// TIA Portal V20 export
Screen "Andon"  1276x673
  ScreenItem "Title_ScreenOverview_X390_Y2" at 9,7 size 1265x44  Type=HmiTextBox
  ScreenItem "permanentareaborderrectangle" at 0,0 size 0x0  Type=HmiRectangle
  ScreenItem "Text box_3" at 346,188 size 590x89  Type=HmiTextBox
  ScreenItem "Title_ScreenOverview_X390_Y2_1" at 9,97 size 84x44  Type=HmiTextBox
  ScreenItem "IO 域_19" at 9,142 size 84x44  Type=HmiIOField
  ScreenItem "Title_ScreenOverview_X390_Y2_5" at 261,97 size 84x44  Type=HmiTextBox
  ScreenItem "IO 域_21" at 261,142 size 84x44  Type=HmiIOField
  ScreenItem "Title_ScreenOverview_X390_Y2_3" at 93,97 size 84x44  Type=HmiTextBox
  ScreenItem "IO 域_5" at 93,142 size 84x44  Type=HmiIOField
  ScreenItem "Title_ScreenOverview_X390_Y2_4" at 177,97 size 84x44  Type=HmiTextBox
  ScreenItem "IO 域_20" at 177,142 size 84x44  Type=HmiIOField
  ScreenItem "Title_ScreenOverview_X390_Y2_6" at 345,97 size 84x44  Type=HmiTextBox
  ScreenItem "IO 域_22" at 345,142 size 84x44  Type=HmiIOField
  ScreenItem "Title_ScreenOverview_X390_Y2_11" at 9,52 size 252x44  Type=HmiTextBox
  ScreenItem "Title_ScreenOverview_X390_Y2_18" at 431,97 size 84x44  Type=HmiTextBox
  ScreenItem "IO 域_42" at 431,142 size 84x44  Type=HmiIOField
  ScreenItem "Title_ScreenOverview_X390_Y2_19" at 683,97 size 84x44  Type=HmiTextBox
  ScreenItem "IO 域_43" at 683,142 size 84x44  Type=HmiIOField
  ScreenItem "Title_ScreenOverview_X390_Y2_20" at 515,97 size 84x44  Type=HmiTextBox
  ScreenItem "IO 域_44" at 515,142 size 84x44  Type=HmiIOField
  ScreenItem "Title_ScreenOverview_X390_Y2_21" at 599,97 size 84x44  Type=HmiTextBox
  ScreenItem "IO 域_45" at 599,142 size 84x44  Type=HmiIOField
  ScreenItem "Title_ScreenOverview_X390_Y2_22" at 767,97 size 84x44  Type=HmiTextBox
  ScreenItem "IO 域_46" at 767,142 size 84x44  Type=HmiIOField
  ScreenItem "Title_ScreenOverview_X390_Y2_23" at 431,52 size 252x44  Type=HmiTextBox
  ScreenItem "Title_ScreenOverview_X390_Y2_25" at 1105,97 size 84x44  Type=HmiTextBox
  ScreenItem "IO 域_48" at 1105,142 size 84x44  Type=HmiIOField
  ScreenItem "Title_ScreenOverview_X390_Y2_28" at 1189,97 size 84x44  Type=HmiTextBox
  ScreenItem "IO 域_51" at 1189,142 size 84x44  Type=HmiIOField
  ScreenItem "Title_ScreenOverview_X390_Y2_29" at 853,52 size 252x44  Type=HmiTextBox
  ScreenItem "Title_ScreenOverview_X390_Y2_7" at 9,188 size 84x44  Type=HmiTextBox
  ScreenItem "IO 域_23" at 9,233 size 84x44  Type=HmiIOField
  ScreenItem "Title_ScreenOverview_X390_Y2_8" at 177,188 size 84x44  Type=HmiTextBox
  ScreenItem "IO 域_24" at 177,233 size 84x44  Type=HmiIOField
  ScreenItem "Text box_32" at 262,278 size 255x96  Type=HmiTextBox
  ScreenItem "Text box_33" at 514,278 size 255x96  Type=HmiTextBox
  ScreenItem "Text box_34" at 764,278 size 255x96  Type=HmiTextBox
  ScreenItem "Text box_35" at 1017,278 size 255x96  Type=HmiTextBox
  ScreenItem "Text box_36" at 10,373 size 255x96  Type=HmiTextBox
  ScreenItem "Text box_37" at 262,373 size 255x96  Type=HmiTextBox
  ScreenItem "Title_ScreenOverview_X390_Y2_38" at 93,188 size 84x44  Type=HmiTextBox
  ScreenItem "IO 域_6" at 93,233 size 84x44  Type=HmiIOField
  ScreenItem "Title_ScreenOverview_X390_Y2_39" at 261,188 size 84x44  Type=HmiTextBox
  ScreenItem "IO 域_7" at 261,233 size 84x44  Type=HmiIOField
  ScreenItem "Title_ScreenOverview_X390_Y2_24" at 853,97 size 84x44  Type=HmiTextBox
  ScreenItem "IO 域_47" at 853,142 size 84x44  Type=HmiIOField
  ScreenItem "Title_ScreenOverview_X390_Y2_26" at 937,97 size 84x44  Type=HmiTextBox
  ScreenItem "IO 域_49" at 937,142 size 84x44  Type=HmiIOField
  ScreenItem "Title_ScreenOverview_X390_Y2_27" at 1021,97 size 84x44  Type=HmiTextBox
  ScreenItem "IO 域_50" at 1021,142 size 84x44  Type=HmiIOField
  ScreenItem "Title_ScreenOverview_X390_Y2_9" at 937,188 size 84x44  Type=HmiTextBox
  ScreenItem "IO 域_8" at 937,233 size 84x44  Type=HmiIOField
  ScreenItem "Title_ScreenOverview_X390_Y2_10" at 1021,188 size 84x44  Type=HmiTextBox
  ScreenItem "IO 域_9" at 1021,233 size 84x44  Type=HmiIOField
  ScreenItem "Title_ScreenOverview_X390_Y2_14" at 1105,188 size 84x44  Type=HmiTextBox
  ScreenItem "IO 域_10" at 1105,233 size 84x44  Type=HmiIOField
  ScreenItem "Move_Legend" at 1182,7 size 90x44  Type=HmiButton
  ScreenItem "Title_ScreenOverview_X390_Y2_17" at 1189,188 size 84x44  Type=HmiTextBox
  ScreenItem "IO 域_11" at 1189,233 size 84x44  Type=HmiIOField
  ScreenItem "IO field_1" at 9,7 size 168x44  Type=HmiIOField
  ScreenItem "Title_ScreenOverview_X390_Y2_13" at 262,52 size 84x44  Type=HmiTextBox
  ScreenItem "IO 域_12" at 346,52 size 84x44  Type=HmiIOField
  ScreenItem "IO 域_13" at 767,52 size 84x44  Type=HmiIOField
  ScreenItem "Title_ScreenOverview_X390_Y2_15" at 683,52 size 84x44  Type=HmiTextBox
  ScreenItem "IO 域_14" at 1188,53 size 84x44  Type=HmiIOField
  ScreenItem "Title_ScreenOverview_X390_Y2_16" at 1104,53 size 84x44  Type=HmiTextBox
  ScreenItem "IO 域_2" at 504,31 size 126x32  Type=HmiIOField
  ScreenItem "Title_ScreenOverview_X390_Y2_31" at 0,31 size 184x32  Type=HmiTextBox
  ScreenItem "IO 域_4" at 185,31 size 126x32  Type=HmiIOField
  ScreenItem "Title_ScreenOverview_X390_Y2_2" at 0,0 size 630x30  Type=HmiTextBox
  ScreenItem "Title_ScreenOverview_X390_Y2_12" at 313,31 size 189x32  Type=HmiTextBox
  ScreenItem "Title_ScreenOverview_X390_Y2_32" at 0,64 size 184x32  Type=HmiTextBox
  ScreenItem "IO 域_3" at 185,64 size 126x32  Type=HmiIOField
  ScreenItem "Title_ScreenOverview_X390_Y2_30" at 313,64 size 189x32  Type=HmiTextBox
  ScreenItem "IO 域_1" at 504,64 size 126x32  Type=HmiIOField
  ScreenItem "IO 域_57" at 1136,31 size 126x32  Type=HmiIOField
  ScreenItem "Title_ScreenOverview_X390_Y2_33" at 632,31 size 184x32  Type=HmiTextBox
  ScreenItem "IO 域_56" at 817,31 size 126x32  Type=HmiIOField
  ScreenItem "Title_ScreenOverview_X390_Y2_34" at 632,0 size 630x30  Type=HmiTextBox
  ScreenItem "Title_ScreenOverview_X390_Y2_35" at 945,31 size 189x32  Type=HmiTextBox
  ScreenItem "Title_ScreenOverview_X390_Y2_36" at 632,64 size 184x32  Type=HmiTextBox
  ScreenItem "IO 域_58" at 817,64 size 126x32  Type=HmiIOField
  ScreenItem "Title_ScreenOverview_X390_Y2_37" at 945,64 size 189x32  Type=HmiTextBox
  ScreenItem "IO 域_59" at 1136,64 size 126x32  Type=HmiIOField
  ScreenItem "IO 域_37" at 504,31 size 126x32  Type=HmiIOField
  ScreenItem "Title_ScreenOverview_X390_Y2_68" at 0,31 size 184x32  Type=HmiTextBox
  ScreenItem "IO 域_53" at 185,31 size 126x32  Type=HmiIOField
  ScreenItem "Title_ScreenOverview_X390_Y2_67" at 0,0 size 630x30  Type=HmiTextBox
  ScreenItem "Title_ScreenOverview_X390_Y2_66" at 313,31 size 189x32  Type=HmiTextBox
  ScreenItem "Title_ScreenOverview_X390_Y2_65" at 0,64 size 184x32  Type=HmiTextBox
  ScreenItem "IO 域_52" at 185,64 size 126x32  Type=HmiIOField
  ScreenItem "Title_ScreenOverview_X390_Y2_64" at 313,64 size 189x32  Type=HmiTextBox
  ScreenItem "IO 域_41" at 504,64 size 126x32  Type=HmiIOField
  ScreenItem "IO 域_40" at 1136,31 size 126x32  Type=HmiIOField
  ScreenItem "Title_ScreenOverview_X390_Y2_63" at 632,31 size 184x32  Type=HmiTextBox
  ScreenItem "IO 域_39" at 817,31 size 126x32  Type=HmiIOField
  ScreenItem "Title_ScreenOverview_X390_Y2_62" at 632,0 size 630x30  Type=HmiTextBox
  ScreenItem "Title_ScreenOverview_X390_Y2_61" at 945,31 size 189x32  Type=HmiTextBox
  ScreenItem "Title_ScreenOverview_X390_Y2_60" at 632,64 size 184x32  Type=HmiTextBox
  ScreenItem "IO 域_38" at 817,64 size 126x32  Type=HmiIOField
  ScreenItem "Title_ScreenOverview_X390_Y2_69" at 945,64 size 189x32  Type=HmiTextBox
  ScreenItem "IO 域_54" at 1136,64 size 126x32  Type=HmiIOField
  ScreenItem "IO 域_15" at 504,31 size 126x32  Type=HmiIOField
  ScreenItem "Title_ScreenOverview_X390_Y2_48" at 0,31 size 184x32  Type=HmiTextBox
  ScreenItem "IO 域_27" at 185,31 size 126x32  Type=HmiIOField
  ScreenItem "Title_ScreenOverview_X390_Y2_47" at 0,0 size 630x30  Type=HmiTextBox
  ScreenItem "Title_ScreenOverview_X390_Y2_46" at 313,31 size 189x32  Type=HmiTextBox
  ScreenItem "Title_ScreenOverview_X390_Y2_45" at 0,64 size 184x32  Type=HmiTextBox
  ScreenItem "IO 域_26" at 185,64 size 126x32  Type=HmiIOField
  ScreenItem "Title_ScreenOverview_X390_Y2_44" at 313,64 size 189x32  Type=HmiTextBox
  ScreenItem "IO 域_25" at 504,64 size 126x32  Type=HmiIOField
  ScreenItem "IO 域_18" at 1136,31 size 126x32  Type=HmiIOField
  ScreenItem "Title_ScreenOverview_X390_Y2_43" at 632,31 size 184x32  Type=HmiTextBox
  ScreenItem "IO 域_17" at 817,31 size 126x32  Type=HmiIOField
  ScreenItem "Title_ScreenOverview_X390_Y2_42" at 632,0 size 630x30  Type=HmiTextBox
  ScreenItem "Title_ScreenOverview_X390_Y2_41" at 945,31 size 189x32  Type=HmiTextBox
  ScreenItem "Title_ScreenOverview_X390_Y2_40" at 632,64 size 184x32  Type=HmiTextBox
  ScreenItem "IO 域_16" at 817,64 size 126x32  Type=HmiIOField
  ScreenItem "Title_ScreenOverview_X390_Y2_49" at 945,64 size 189x32  Type=HmiTextBox
  ScreenItem "IO 域_28" at 1136,64 size 126x32  Type=HmiIOField
  ScreenItem "IO 域_29" at 504,31 size 126x32  Type=HmiIOField
  ScreenItem "Title_ScreenOverview_X390_Y2_58" at 0,31 size 184x32  Type=HmiTextBox
  ScreenItem "IO 域_35" at 185,31 size 126x32  Type=HmiIOField
  ScreenItem "Title_ScreenOverview_X390_Y2_57" at 0,0 size 630x30  Type=HmiTextBox
  ScreenItem "Title_ScreenOverview_X390_Y2_56" at 313,31 size 189x32  Type=HmiTextBox
  ScreenItem "Title_ScreenOverview_X390_Y2_55" at 0,64 size 184x32  Type=HmiTextBox
  ScreenItem "IO 域_34" at 185,64 size 126x32  Type=HmiIOField
  ScreenItem "Title_ScreenOverview_X390_Y2_54" at 313,64 size 189x32  Type=HmiTextBox
  ScreenItem "IO 域_33" at 504,64 size 126x32  Type=HmiIOField
  ScreenItem "IO 域_32" at 1136,31 size 126x32  Type=HmiIOField
  ScreenItem "Title_ScreenOverview_X390_Y2_53" at 632,31 size 184x32  Type=HmiTextBox
  ScreenItem "IO 域_31" at 817,31 size 126x32  Type=HmiIOField
  ScreenItem "Title_ScreenOverview_X390_Y2_52" at 632,0 size 630x30  Type=HmiTextBox
  ScreenItem "Title_ScreenOverview_X390_Y2_51" at 945,31 size 189x32  Type=HmiTextBox
  ScreenItem "Title_ScreenOverview_X390_Y2_50" at 632,64 size 184x32  Type=HmiTextBox
  ScreenItem "IO 域_30" at 817,64 size 126x32  Type=HmiIOField
  ScreenItem "Title_ScreenOverview_X390_Y2_59" at 945,64 size 189x32  Type=HmiTextBox
  ScreenItem "IO 域_36" at 1136,64 size 126x32  Type=HmiIOField
  ScreenItem "Text box_1" at 514,373 size 255x96  Type=HmiTextBox
  ScreenItem "Text box_2" at 10,278 size 255x96  Type=HmiTextBox
  ScreenItem "Text box_4" at 764,373 size 255x96  Type=HmiTextBox
  ScreenItem "Text box_5" at 1017,373 size 255x96  Type=HmiTextBox
  ScreenItem "Text box_6" at 10,469 size 255x96  Type=HmiTextBox
  ScreenItem "Text box_7" at 262,469 size 255x96  Type=HmiTextBox
  ScreenItem "Text box_8" at 514,469 size 255x96  Type=HmiTextBox
  ScreenItem "Text box_9" at 764,469 size 255x96  Type=HmiTextBox
  ScreenItem "IO 域_55" at 504,31 size 126x32  Type=HmiIOField
  ScreenItem "Title_ScreenOverview_X390_Y2_78" at 0,31 size 184x32  Type=HmiTextBox
  ScreenItem "IO 域_65" at 185,31 size 126x32  Type=HmiIOField
  ScreenItem "Title_ScreenOverview_X390_Y2_77" at 0,0 size 630x30  Type=HmiTextBox
  ScreenItem "Title_ScreenOverview_X390_Y2_76" at 313,31 size 189x32  Type=HmiTextBox
  ScreenItem "Title_ScreenOverview_X390_Y2_75" at 0,64 size 184x32  Type=HmiTextBox
  ScreenItem "IO 域_64" at 185,64 size 126x32  Type=HmiIOField
  ScreenItem "Title_ScreenOverview_X390_Y2_74" at 313,64 size 189x32  Type=HmiTextBox
  ScreenItem "IO 域_63" at 504,64 size 126x32  Type=HmiIOField
  ScreenItem "IO 域_62" at 1136,31 size 126x32  Type=HmiIOField
  ScreenItem "Title_ScreenOverview_X390_Y2_73" at 632,31 size 184x32  Type=HmiTextBox
  ScreenItem "IO 域_61" at 817,31 size 126x32  Type=HmiIOField
  ScreenItem "Title_ScreenOverview_X390_Y2_72" at 632,0 size 630x30  Type=HmiTextBox
  ScreenItem "Title_ScreenOverview_X390_Y2_71" at 945,31 size 189x32  Type=HmiTextBox
  ScreenItem "Title_ScreenOverview_X390_Y2_70" at 632,64 size 184x32  Type=HmiTextBox
  ScreenItem "IO 域_60" at 817,64 size 126x32  Type=HmiIOField
  ScreenItem "Title_ScreenOverview_X390_Y2_79" at 945,64 size 189x32  Type=HmiTextBox
  ScreenItem "IO 域_66" at 1136,64 size 126x32  Type=HmiIOField
  ScreenItem "IO 域_67" at 504,31 size 126x32  Type=HmiIOField
  ScreenItem "Title_ScreenOverview_X390_Y2_88" at 0,31 size 184x32  Type=HmiTextBox
  ScreenItem "IO 域_73" at 185,31 size 126x32  Type=HmiIOField
  ScreenItem "Title_ScreenOverview_X390_Y2_89" at 0,0 size 630x30  Type=HmiTextBox
  ScreenItem "Title_ScreenOverview_X390_Y2_87" at 313,31 size 189x32  Type=HmiTextBox
  ScreenItem "Title_ScreenOverview_X390_Y2_86" at 0,64 size 184x32  Type=HmiTextBox
  ScreenItem "IO 域_72" at 185,64 size 126x32  Type=HmiIOField
  ScreenItem "Title_ScreenOverview_X390_Y2_85" at 313,64 size 189x32  Type=HmiTextBox
  ScreenItem "IO 域_71" at 504,64 size 126x32  Type=HmiIOField
  ScreenItem "IO 域_70" at 1136,31 size 126x32  Type=HmiIOField
  ScreenItem "Title_ScreenOverview_X390_Y2_84" at 632,31 size 184x32  Type=HmiTextBox
  ScreenItem "IO 域_69" at 817,31 size 126x32  Type=HmiIOField
  ScreenItem "Title_ScreenOverview_X390_Y2_83" at 632,0 size 630x30  Type=HmiTextBox
  ScreenItem "Title_ScreenOverview_X390_Y2_82" at 945,31 size 189x32  Type=HmiTextBox
  ScreenItem "Title_ScreenOverview_X390_Y2_81" at 632,64 size 184x32  Type=HmiTextBox
  ScreenItem "IO 域_68" at 817,64 size 126x32  Type=HmiIOField
  ScreenItem "Title_ScreenOverview_X390_Y2_80" at 945,64 size 189x32  Type=HmiTextBox
  ScreenItem "IO 域_74" at 1136,64 size 126x32  Type=HmiIOField
  ScreenItem "IO 域_75" at 504,31 size 126x32  Type=HmiIOField
  ScreenItem "Title_ScreenOverview_X390_Y2_98" at 0,31 size 184x32  Type=HmiTextBox
  ScreenItem "IO 域_81" at 185,31 size 126x32  Type=HmiIOField
  ScreenItem "Title_ScreenOverview_X390_Y2_99" at 0,0 size 630x30  Type=HmiTextBox
  ScreenItem "Title_ScreenOverview_X390_Y2_97" at 313,31 size 189x32  Type=HmiTextBox
  ScreenItem "Title_ScreenOverview_X390_Y2_96" at 0,64 size 184x32  Type=HmiTextBox
  ScreenItem "IO 域_80" at 185,64 size 126x32  Type=HmiIOField
  ScreenItem "Title_ScreenOverview_X390_Y2_95" at 313,64 size 189x32  Type=HmiTextBox
  ScreenItem "IO 域_79" at 504,64 size 126x32  Type=HmiIOField
  ScreenItem "IO 域_78" at 1136,31 size 126x32  Type=HmiIOField
  ScreenItem "Title_ScreenOverview_X390_Y2_94" at 632,31 size 184x32  Type=HmiTextBox
  ScreenItem "IO 域_77" at 817,31 size 126x32  Type=HmiIOField
  ScreenItem "Title_ScreenOverview_X390_Y2_93" at 632,0 size 630x30  Type=HmiTextBox
  ScreenItem "Title_ScreenOverview_X390_Y2_92" at 945,31 size 189x32  Type=HmiTextBox
  ScreenItem "Title_ScreenOverview_X390_Y2_91" at 632,64 size 184x32  Type=HmiTextBox
  ScreenItem "IO 域_76" at 817,64 size 126x32  Type=HmiIOField
  ScreenItem "Title_ScreenOverview_X390_Y2_90" at 945,64 size 189x32  Type=HmiTextBox
  ScreenItem "IO 域_82" at 1136,64 size 126x32  Type=HmiIOField
  ScreenItem "Rectangle_36" at 297,0 size 115x81  Type=HmiRectangle
  ScreenItem "Text_38" at 297,15 size 115x51  Type=HmiText
  ScreenItem "Rectangle_37" at 0,87 size 144x46  Type=HmiRectangle
  ScreenItem "Text_39" at 5,90 size 133x38  Type=HmiText
  ScreenItem "Rectangle_38" at 0,0 size 144x46  Type=HmiRectangle
  ScreenItem "Text_40" at 8,10 size 133x27  Type=HmiText
  ScreenItem "Rectangle_39" at 143,87 size 155x46  Type=HmiRectangle
  ScreenItem "Text_41" at 189,97 size 64x28  Type=HmiText
  ScreenItem "Rectangle_40" at 143,0 size 155x46  Type=HmiRectangle
  ScreenItem "Text_42" at 183,9 size 76x32  Type=HmiText
  ScreenItem "Rectangle_31" at 297,0 size 115x81  Type=HmiRectangle
  ScreenItem "Text_33" at 297,15 size 115x51  Type=HmiText
  ScreenItem "Rectangle_32" at 0,87 size 144x46  Type=HmiRectangle
  ScreenItem "Text_34" at 5,90 size 133x38  Type=HmiText
  ScreenItem "Rectangle_33" at 0,0 size 144x46  Type=HmiRectangle
  ScreenItem "Text_35" at 8,10 size 133x27  Type=HmiText
  ScreenItem "Rectangle_34" at 143,87 size 155x46  Type=HmiRectangle
  ScreenItem "Text_36" at 189,97 size 64x28  Type=HmiText
  ScreenItem "Rectangle_35" at 143,0 size 155x46  Type=HmiRectangle
  ScreenItem "Text_37" at 183,9 size 76x32  Type=HmiText
